(* IEC 61131-3 sources: verifaps-lib/stvs/src/test/resources/edu/kit/iti/formal/stvs/testSets/valid_1, 1 file *)

(* ---- code_valid_1.st ---- *)
TYPE
  enumD : (literalOne, literalTwo);
END_TYPE

PROGRAM constantprogram
  VAR_INPUT
    A : INT;
    B : BOOL;
  END_VAR

  VAR_OUTPUT
    C : INT;
    D : enumD;
  END_VAR

  C := 52;
END_PROGRAM
